Yaskawa INFORM job: SPLITTE3.JBI

/JOB
//NAME SPLITTE3
//POS
///NPOS 15,0,0,0,0,0
///TOOL 1
///POSTYPE BASE
///RECTAN
///RCONF 0,0,0,0,0,0,0,0
C00000=661.027,82.386,686.221,-67.04,7.80,-111.79
C00001=674.300,134.999,685.980,-66.22,8.38,-107.67
C00002=661.027,82.386,686.221,-67.04,7.80,-111.79
C00003=674.300,134.999,685.980,-66.22,8.38,-107.67
C00004=661.027,82.386,686.221,-67.04,7.80,-111.79
C00005=674.300,134.999,685.980,-66.22,8.38,-107.67
C00006=661.027,82.386,686.221,-67.04,7.80,-111.79
C00007=674.300,134.999,685.980,-66.22,8.38,-107.67
C00008=661.027,82.386,686.221,-67.04,7.80,-111.79
C00009=674.300,134.999,685.980,-66.22,8.38,-107.67
C00010=661.027,82.386,686.221,-67.04,7.80,-111.79
C00011=674.300,134.999,685.980,-66.22,8.38,-107.67
C00012=661.027,82.386,686.221,-67.04,7.80,-111.79
C00013=674.300,134.999,685.980,-66.22,8.38,-107.67
C00014=661.027,82.386,686.221,-67.04,7.80,-111.79
//INST
///DATE 2026/10/26 01:19
///COMM Generated using RoboDK
///ATTR SC,RW,RJ
///GROUP1 RB1
NOP
MOVL C00000 V=200.0
MOVL C00001 V=200.0
MOVL C00002 V=200.0
MOVL C00003 V=200.0
MOVL C00004 V=200.0
MOVL C00005 V=200.0
MOVL C00006 V=200.0
MOVL C00007 V=200.0
MOVL C00008 V=200.0
MOVL C00009 V=200.0
MOVL C00010 V=200.0
MOVL C00011 V=200.0
MOVL C00012 V=200.0
MOVL C00013 V=200.0
MOVL C00014 V=200.0
END
